RoboDK station: Car_Painting_Cell_v2.rdk

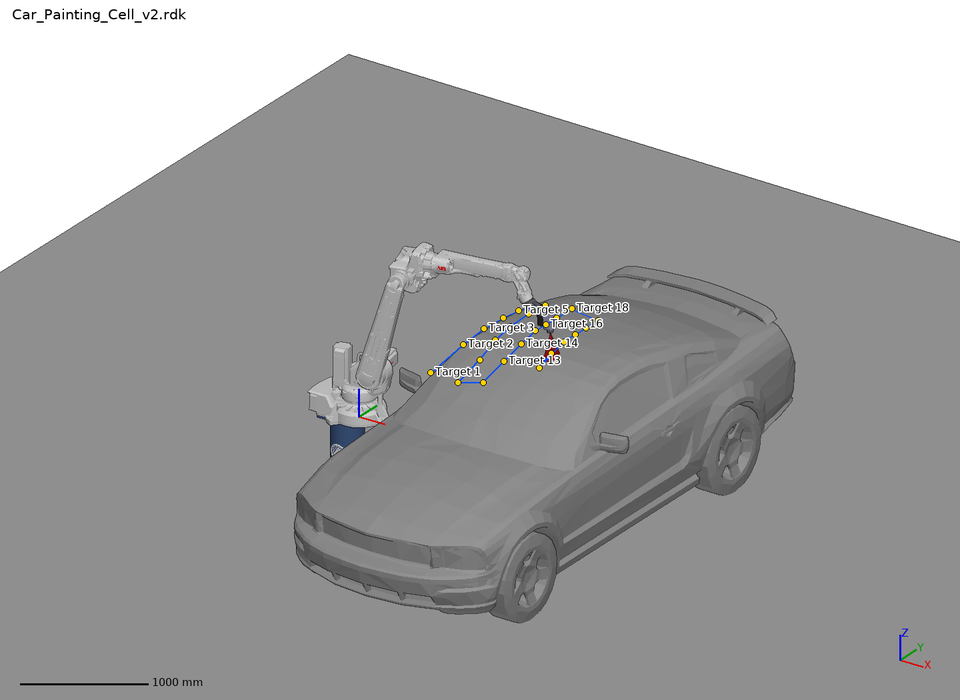
[picture v0: the station drawn from its stored meshes, robots at their saved joint values, targets as dots, program paths as lines]
Station Car_Painting_Cell_v2 (saved by RoboDK 6.1.1). Poses are relative to the parent item; angles as X-Y-Z fixed-axis rotations.
  - object 78256 at (0, 0, 0) mm, size 2178.4 x 4892.4 x 1442.1 mm, geometry from 78256.obj
  - object Floor at (0, 0, 0) mm, size 12000 x 12000 x 0 mm, geometry from Floor.sld
  - frame ABB IRB 2600ID-8/2.00 Base at (-1520, -250, 600) mm
    - robot ABB IRB 2600ID-8/2.00: 6 axes, payload 8 kg, reach 2000 mm, repeatability 0.023 mm, weight 276 kg
        modified DH rows (alpha deg, a mm, theta deg, d mm): 0, 0, 0, 445; -90, 150, -90, 0; 0, 900, 0, 0; -90, 150, 0, 938; 90, 0, 0, 0; -90, 0, 180, 200
        joint limits [-180, -95, -180, -175, -120, -400] to [180, 155, 75, 175, 120, 400]; home [0, 0, 0, 0, 0, 0]; saved at [11.695, 15.5, -14.491, -0.903, 57.055, 7.158]
      - tool Generic Paint Sprayer, TCP at (50, 0, 450) mm, rotated rx 0 ry 30 rz 0 deg, size 277.6 x 203.2 x 501.7 mm
    - target Target 1 (Cartesian target) at (786.75, -147.83, 660.16) mm, rotated rx 162.25 ry 7.56 rz 171.38 deg; joints [-33.508, -42.216, 47.281, 34.8, 59.888, -32.291] of ABB IRB 2600ID-8/2.00
    - target Target 2 (Cartesian target) at (845.19, 209.11, 778.74) mm, rotated rx 170.39 ry 7.35 rz 175.51 deg; joints [15.978, -39.932, 37.942, -5.407, 53.846, 24.142] of ABB IRB 2600ID-8/2.00
    - target Target 3 (Cartesian target) at (850.9, 479.97, 809.5) mm, rotated rx 179.56 ry 8.38 rz -177.95 deg; joints [43.521, -27.96, 30.387, -28.018, 59.845, 49.81] of ABB IRB 2600ID-8/2.00
    - target Target 4 (Cartesian target) at (851.43, 746.82, 799.82) mm, rotated rx -174.47 ry 15.36 rz -170.53 deg; joints [60.093, -16.443, 26.657, -44.197, 59.731, 66.095] of ABB IRB 2600ID-8/2.00
    - target Target 5 (Cartesian target) at (802.88, 1027.63, 735.48) mm, rotated rx -164.76 ry 30.87 rz -166.22 deg; joints [76.691, 1.156, 24.253, -68.858, 68.439, 93.616] of ABB IRB 2600ID-8/2.00
    - target Target 6 (Cartesian target) at (964.94, 1158.15, 773.42) mm, rotated rx -170.29 ry 3.53 rz -171.47 deg; joints [62.224, 17.274, -10.002, -33.97, 71.871, 59.088] of ABB IRB 2600ID-8/2.00
    - target Target 7 (Cartesian target) at (990.36, 891.41, 812.91) mm, rotated rx -172.68 ry 3.03 rz -171.54 deg; joints [53.897, 2.48, 4.423, -30.544, 66.343, 51.971] of ABB IRB 2600ID-8/2.00
    - target Target 8 (Cartesian target) at (1035.85, 583.51, 840.52) mm, rotated rx -177.89 ry 1.87 rz -171.58 deg; joints [37.338, -10.949, 14.603, -19.084, 60.005, 34.107] of ABB IRB 2600ID-8/2.00
    - target Target 9 (Cartesian target) at (1071.58, 321.15, 835.07) mm, rotated rx 179.21 ry 2.98 rz -171.6 deg; joints [19.295, -18.39, 20.918, -6.386, 55.026, 13.223] of ABB IRB 2600ID-8/2.00
    - target Target 10 (Cartesian target) at (1112.71, 50.86, 784.62) mm, rotated rx 170.71 ry 4.64 rz -171.87 deg; joints [-6.364, -18.947, 25.383, 20.329, 52.975, -20.23] of ABB IRB 2600ID-8/2.00
    - target Target 11 (Cartesian target) at (1084.41, -204.31, 682.79) mm, rotated rx 162.98 ry 8.07 rz -172.92 deg; joints [-29.187, -15.026, 31.029, 42.116, 57.57, -50.949] of ABB IRB 2600ID-8/2.00
    - target Target 12 (Cartesian target) at (1286.21, -152.58, 718.35) mm, rotated rx 163.83 ry 3.37 rz -178.07 deg; joints [-18.486, -4.211, 17.952, 31.68, 52.597, -30.766] of ABB IRB 2600ID-8/2.00
    - target Target 13 (Cartesian target) at (1307.72, 101.1, 804.5) mm, rotated rx 170.22 ry 3.47 rz -178.83 deg; joints [-0.3, -6.762, 14.218, 12.231, 49.548, -4.318] of ABB IRB 2600ID-8/2.00
    - target Target 14 (Cartesian target) at (1303.7, 348.12, 858.06) mm, rotated rx -177.91 ry 1.89 rz -172.09 deg; joints [18.112, -2.578, 6.113, -8.696, 55.554, 12.62] of ABB IRB 2600ID-8/2.00
    - target Target 15 (Cartesian target) at (1288.42, 553.54, 885.8) mm, rotated rx -171.33 ry 2.81 rz -171.95 deg; joints [31.671, 2.872, -0.351, -22.558, 61.326, 27.799] of ABB IRB 2600ID-8/2.00
    - target Target 16 (Cartesian target) at (1262.24, 740.76, 857.97) mm, rotated rx -171.13 ry 0.58 rz -172.3 deg; joints [39.375, 9.876, -7.096, -24.588, 66.198, 35.173] of ABB IRB 2600ID-8/2.00
    - target Target 17 (Cartesian target) at (1234.75, 919.61, 834.98) mm, rotated rx -176.98 ry 0.53 rz -172.31 deg; joints [43.946, 14.114, -11.168, -21.888, 64.759, 40.95] of ABB IRB 2600ID-8/2.00
    - target Target 18 (Cartesian target) at (1206.03, 1172.88, 805.97) mm, rotated rx -172.14 ry 2.41 rz -172.62 deg; joints [53.666, 27.49, -26.431, -29.443, 72.541, 49.22] of ABB IRB 2600ID-8/2.00
    - target Target 19 (Cartesian target) at (1512.91, 1087.25, 824.86) mm, rotated rx -177.34 ry 2.14 rz -175.71 deg; joints [42.099, 38.739, -45.176, -22.018, 72.644, 39.315] of ABB IRB 2600ID-8/2.00
    - target Target 21 (Cartesian target) at (1544.21, 733.41, 849.84) mm, rotated rx -174.5 ry 0.23 rz -173.93 deg; joints [31.162, 25.245, -26.767, -18.337, 66.559, 27.232] of ABB IRB 2600ID-8/2.00
    - target Target 20 (Cartesian target) at (1532.94, 899.54, 837.3) mm, rotated rx 178.9 ry -0.74 rz -175.83 deg; joints [34.565, 30.245, -33.698, -14.564, 67.873, 33.133] of ABB IRB 2600ID-8/2.00
    - target Target 22 (Cartesian target) at (1567.73, 545.31, 871.98) mm, rotated rx -171.81 ry 0.14 rz -172.36 deg; joints [24.84, 20.894, -21.957, -17.13, 64.706, 18.728] of ABB IRB 2600ID-8/2.00
    - target Target 23 (Cartesian target) at (1623.15, 130.83, 824.97) mm, rotated rx 169.94 ry 6.74 rz -175.3 deg; joints [-0.004, 11.93, -5.331, 15.592, 48.019, -9.331] of ABB IRB 2600ID-8/2.00
    - target Target 24 (Cartesian target) at (1599.3, 329.18, 868.05) mm, rotated rx 177.15 ry 1.8 rz -174.46 deg; joints [11.75, 15.529, -14.549, -0.969, 57.113, 7.221] of ABB IRB 2600ID-8/2.00
  - object Pedestal H24in (Type 1) at (-1640, -240, 0) mm, size 400 x 400 x 609.6 mm, geometry from Pedestal-H24in-Type-1.sld
  - program Prog1 (26 instructions, listed below)
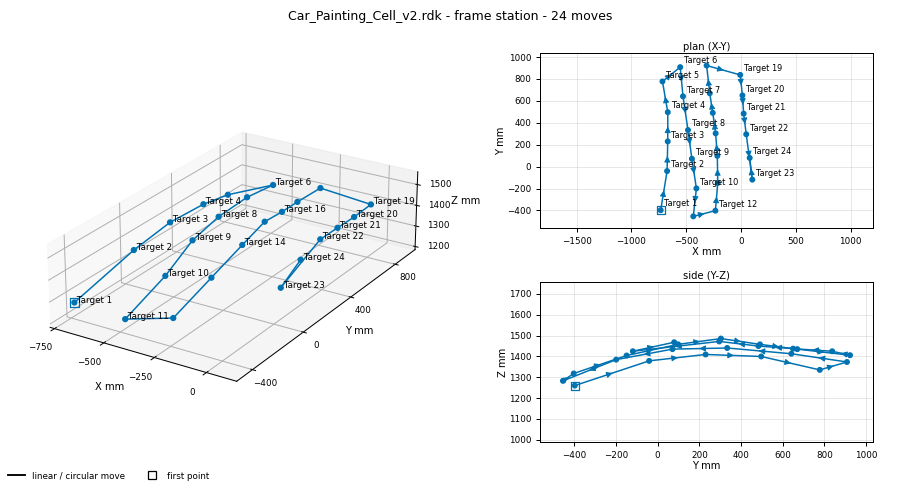
[picture p0: tool path of Car_Painting_Cell_v2.rdk in frame station, 24 of 24 moves have a stored position in this frame; points joined in program order, loops and branches not executed]

--- program Prog1 (robot ABB IRB 2600ID-8/2.00) ---
  Set Ref.: ABB IRB 2600ID-8/2.00 Base
  Set Tool: Generic Paint Sprayer
  MoveJ (Target 1)
  MoveL (Target 2)
  MoveL (Target 3)
  MoveL (Target 4)
  MoveL (Target 5)
  MoveL (Target 6)
  MoveL (Target 7)
  MoveL (Target 8)
  MoveL (Target 9)
  MoveL (Target 10)
  MoveL (Target 11)
  MoveL (Target 12)
  MoveL (Target 13)
  MoveL (Target 14)
  MoveL (Target 15)
  MoveL (Target 16)
  MoveL (Target 17)
  MoveL (Target 18)
  MoveL (Target 19)
  MoveL (Target 20)
  MoveL (Target 21)
  MoveL (Target 22)
  MoveL (Target 23)
  MoveL (Target 24)
